Fanuc KAREL source: ka00130.KL

-- PROVISIONAL review KL for V1013-1; original PC SHA256 8e545cfdbf0790b4862ca504e5f6dad9aed0f27cda0d552aa24a88a868bf71e7
-- Incomplete behavior may be omitted. Consult companion uncertainty JSON. Do not deploy.
PROGRAM KA00130
%NOLOCKGROUP
-- UNRESOLVED_DECL SRC type=002018
-- UNRESOLVED_DECL DST type=00001c
BEGIN
  -- UNRESOLVED_PC offsets 5-19; opcodes 2E,22,9D,33,B2
  -- UNRESOLVED_PC offsets 24-39; opcodes 22,9D,33,B1,23
  -- UNRESOLVED_PC offsets 44-48; opcodes 7F
END KA00130
